(* IEC 61131-3 sources: repo_PLC_code_eval/dataset/2021-8-20/F03_气缸操作, 3 files *)

(* ---- FB_气缸延时.st ---- *)
FUNCTION_BLOCK FB_气缸延时
VAR_INPUT
	Clinyder: BOOL;
	OpenDelayTime: REAL;
	CloseDelayTime: REAL;
	OpenSensor: BOOL;
	CloseSensor: BOOL;
END_VAR
VAR_OUTPUT
	OpenDelay: BOOL;
	CloseDelay: BOOL;
END_VAR
VAR
	TON0: TON;
	TON1: TON;
END_VAR

TON0(IN:= Clinyder , PT:= REAL_TO_TIME(OpenDelayTime*1000), Q=> , ET=> );
TON1(IN:= NOT Clinyder , PT:= REAL_TO_TIME(CloseDelayTime*1000), Q=> , ET=> );

IF TON0.Q THEN
	OpenDelay:=TRUE;
	ELSE
	OpenDelay:=FALSE;
END_IF

IF TON1.Q THEN
	CloseDelay:=TRUE;
	ELSE
	CloseDelay:=FALSE;
END_IF

(* ---- FB_气缸手动111111.st ---- *)
FUNCTION_BLOCK FB_气缸手动
VAR_INPUT
	Excute: BOOL;
END_VAR
VAR_OUTPUT
	Out: BOOL;
END_VAR
VAR
	R_TRIG_0: R_TRIG;
	F_TRIG_0: F_TRIG;
END_VAR

(* ---- FB_气缸操作块1111111.st ---- *)
FUNCTION_BLOCK FB_气缸操作块
VAR_INPUT
	CheckTime: TIME := T#3S;
	OpenSensor: BOOL;
	CloseSensor: BOOL;

	OpenSensorCheck: BOOL;
	CloseSensorCheck: BOOL;

	OpenDelayTime: REAL;
	CloseDelayTime: REAL;

	Cylinder: BOOL;
END_VAR

VAR_OUTPUT
	Q_CylinderError1: BOOL;
	Q_CylinderError2: BOOL;
	OpenDelay: BOOL;
	CloseDelay: BOOL;
END_VAR
VAR
	Delay1: TON;
	Delay2: TON;
	TON0: TON;
	TON1: TON;
END_VAR
